FUNCTION_BLOCK FB_Conveyor
VAR_INPUT
	
	Start			:	BOOL;
	Stop			:	BOOL;
	EmergencyStop	:	BOOL;
	Reset			:	BOOL;
	
	AutoMode      	:	BOOL;
	SensorEntry   	: 	BOOL;
    SensorExit    	: 	BOOL;
	
	Mode	:	E_ConveyorMode;
	
END_VAR
VAR_OUTPUT
	
	Motor 		: BOOL;
	GreenLamp 	: BOOL;
	RedLamp 	: BOOL;
	FaultLamp	: BOOL;
	
	FaultCode : E_FaultCode := E_FaultCode.FC_NONE;
	
	
	
END_VAR
VAR
	
   
   
	
	State 	: 	E_ConveyorState ;
	
	
	ModeChanged 	: BOOL;
    PreviousMode 	: E_ConveyorMode;

  
	
	TimerPart		:	TON;
	ExitTrigger		:	R_TRIG;
	EntryTrigger 	: 	R_TRIG;
	Counter 		: 	UDINT := 0;
	
	InterlockOK 	: 	BOOL;
	
	
	
	
	
END_VAR

TimerPart(
    	IN := (Mode = E_ConveyorMode.AUTO)
          	AND 
				(State = E_ConveyorState.WAIT_EXIT),
    	PT := T#10S
	);
ExitTrigger(CLK := SensorExit);	
EntryTrigger(CLK := SensorEntry);
ModeChanged := Mode <> PreviousMode;

IF NOT HandleFaults() THEN
    IF NOT HandleModeChange() THEN
        IF Mode = E_ConveyorMode.AUTO THEN
            RunAuto();

        ELSIF Mode = E_ConveyorMode.MANUAL THEN
            RunManual();
        END_IF
    END_IF
END_IF

UpdateOutputs();

METHOD HandleFaults : BOOL
VAR_INPUT
END_VAR

VAR
END_VAR
HandleFaults := FALSE;

IF EmergencyStop THEN
    State := E_ConveyorState.FAULT;
    FaultCode := E_FaultCode.FC_EMERGENCY_STOP;
    HandleFaults := TRUE;

ELSIF Reset AND State = E_ConveyorState.FAULT THEN
    State := E_ConveyorState.IDLE;
    FaultCode := E_FaultCode.FC_NONE;
    HandleFaults := TRUE;

ELSIF State = E_ConveyorState.FAULT THEN
    HandleFaults := TRUE;
END_IF
END_METHOD

METHOD HandleModeChange : BOOL
VAR_INPUT
END_VAR
HandleModeChange := FALSE;

IF ModeChanged THEN
    IF State <> E_ConveyorState.FAULT THEN
        State := E_ConveyorState.IDLE;
    END_IF

    HandleModeChange := TRUE;
END_IF
END_METHOD

METHOD RunAuto
VAR_INPUT
END_VAR
IF SensorExit THEN
    InterlockOK := FALSE;
ELSE
    InterlockOK := TRUE;
END_IF

CASE State OF

    E_ConveyorState.IDLE:
        IF Start AND InterlockOK THEN
            State := E_ConveyorState.RUNNING;
        END_IF

    E_ConveyorState.RUNNING:
        IF EntryTrigger.Q THEN
            State := E_ConveyorState.WAIT_EXIT;
        ELSIF Stop THEN
            State := E_ConveyorState.IDLE;
        END_IF

    E_ConveyorState.WAIT_EXIT:
        IF TimerPart.Q THEN
            State := E_ConveyorState.FAULT;
            FaultCode := E_FaultCode.FC_EXIT_TIMEOUT;
        ELSIF ExitTrigger.Q THEN
            State := E_ConveyorState.RUNNING;
            Counter := Counter + 1;
        ELSIF Stop THEN
            State := E_ConveyorState.IDLE;
        END_IF

END_CASE
END_METHOD

METHOD RunManual
VAR_INPUT
END_VAR
IF State <> E_ConveyorState.FAULT THEN
    IF Start THEN
        State := E_ConveyorState.RUNNING;
    ELSE
        State := E_ConveyorState.IDLE;
    END_IF
END_IF
END_METHOD

METHOD UpdateOutputs
VAR_INPUT
END_VAR
Motor := (State = E_ConveyorState.RUNNING)
      OR (State = E_ConveyorState.WAIT_EXIT);

GreenLamp := Motor;
RedLamp := State = E_ConveyorState.IDLE;
FaultLamp := State = E_ConveyorState.FAULT;
END_METHOD

END_FUNCTION_BLOCK

(* stored: Version 1.1.0.1, ProductVersion 3.1.4026.21
   POU FB_Conveyor: Id {e691a8aa-df53-4498-ae74-d15bcd0b3190}, SpecialFunc None
   Method HandleFaults: Id {0142073b-7014-404b-b3cf-64a9e958afe6}
   Method HandleModeChange: Id {61773f67-d62d-4761-8a96-fe95c768418b}
   Method RunAuto: Id {1694a31d-b738-4af3-b469-e300ec7d2e2d}
   Method RunManual: Id {d7dffffb-616f-4be3-b62f-b75890a221ae}
   Method UpdateOutputs: Id {15c67a64-11fb-4727-b413-a2890330b365} *)
